// TIA Portal V19 export
TYPE "ST_Power"
   STRUCT
      Enable : Bool;
      Enabled : Bool;
      Error : Bool;
      ErrorID : Word;
   END_STRUCT;
END_TYPE
